TYPE ST_YARD_CTRL :
STRUCT
  Cmd                     : E_INSTANCE_CMD;
END_STRUCT
END_TYPE

(* stored: Version 1.1.0.1
   DUT ST_YARD_CTRL: Id {616260e5-de48-46b7-a15a-8d70e24db40b} *)
